NAMESPACE TiaMcp_UnitA.Alternate
DATA_BLOCK "TgpNamespace_GlobalTonr"
{ S7_Optimized_Access := 'TRUE' }
VERSION : 0.1
"IEC_TIMER"
BEGIN
END_DATA_BLOCK

END_NAMESPACE
